{attribute 'qualified_only'}
VAR_GLOBAL CONSTANT
	MAX_SCAN_POINTS : UINT := 1024;
	SIMULATOR_PROTOCOL_VERSION : UDINT := 2;
	SIMULATOR_TIMEOUT_IN_CYCLES : UDINT := 20;
	LIDAR_TIMEOUT_IN_MS : TIME := T#400MS;
	SIMULATOR_NOT_CONNECTED_ERROR_ID : UDINT := 1001;
	LIDAR_TIMEOUT_ERROR_ID : UDINT := 2001;
	AXIS_NOT_LINKED_ERROR_ID : UDINT := 3001;
END_VAR

(* stored: Version 1.1.0.1, ProductVersion 3.1.4026.12
   GVL Constants: Id {f17f1f5b-9325-54fe-af2c-f89a3e9a99bf} *)
